(* IEC 61131-3 sources: Versio-VersionControlSystem/fixtures/projects/MachineWithMembers/Device/Plc Logic/Application/Pumps, 1 file *)

(* ---- FB_Pump.st ---- *)
FUNCTION_BLOCK FB_Pump
VAR_INPUT
	enable : BOOL;
END_VAR
VAR_OUTPUT
	running : BOOL;
END_VAR
VAR
	speed : INT;
END_VAR

// --- BEGIN IMPLEMENTATION ---

running := enable;
